Fanuc KAREL source: ka00118.KL

-- PROVISIONAL review KL for V1013-1; original PC SHA256 52d5c9f54aed98fa3839e2e2026405d7d35df101179b3f8a5da9c50ed1834722
-- Incomplete behavior may be omitted. Consult companion uncertainty JSON. Do not deploy.
PROGRAM KA00118
%NOLOCKGROUP
-- UNRESOLVED_DECL SRC type=00001c
-- UNRESOLVED_DECL DST type=00001c
BEGIN
  -- UNRESOLVED_PC offsets 5-15; opcodes 9D,22,A5
  -- UNRESOLVED_PC offsets 20-32; opcodes 21,23
  -- UNRESOLVED_PC offsets 37-41; opcodes 7F
END KA00118
